// TIA Portal V20 export
DATA_BLOCK "DB_ALARM"   // DB100
{ S7_Optimized_Access := 'FALSE' }
// stored: AutoNumber false
   VAR
      ALARM : Struct
         ALARM_GLOBAL : Bool;   // globální alarm
         HERMA_ERROR : Bool;
         ALARM_2 : Bool;
         ALARM_3 : Bool;
         ALARM_4 : Bool;
         ALARM_5 : Bool;
         air : Bool;   // nedostatečný tlak vzduchu
         ALARM_7 : Bool;
         ALARM_8 : Bool;
         ALARM_9 : Bool;
         ALARM_10 : Bool;
         ALARM_11 : Bool;
         ALARM_12 : Bool;
         ALARM_13 : Bool;
         ALARM_14 : Bool;
         vypadek_safety_karty : Bool;
      END_STRUCT;
      WRONG : Struct
         NENI_INICIALIZACE : Bool;
         WRONG_global : Bool;
         dvere_L_tevreny : Bool;
         dvere_P_otevreny : Bool;
         WRONG_4 : Bool;
         WRONG_5 : Bool;
         WRONG_6 : Bool;
         WRONG_7 : Bool;
         WRONG_8 : Bool;
         WRONG_9 : Bool;
         WRONG_10 : Bool;
         WRONG_11 : Bool;
         WRONG_12 : Bool;
         WRONG_13 : Bool;
         rop_glob_warning : Bool;
         rop_active_autocale : Bool;
      END_STRUCT;
      OP0 : Struct
         ALARM : Struct
            DOOR_ERROR : Bool;
            ALARM_1 : Bool;
            ALARM_2 : Bool;
            ALARM_3 : Bool;
            ALARM_4 : Bool;
            ALARM_5 : Bool;
            ALARM_6 : Bool;
            ALARM_7 : Bool;
            ALARM_8 : Bool;
            ALARM_9 : Bool;
            ALARM_10 : Bool;
            ALARM_11 : Bool;
            ALARM_12 : Bool;
            ALARM_13 : Bool;
            ALARM_14 : Bool;
            ALARM_15 : Bool;
         END_STRUCT;
         WRONG : Struct
            WRONG_0 : Bool;
            WRONG_1 : Bool;
            WRONG_2 : Bool;
            WRONG_3 : Bool;
            WRONG_4 : Bool;
            WRONG_5 : Bool;
            WRONG_6 : Bool;
            WRONG_7 : Bool;
            WRONG_8 : Bool;
            WRONG_9 : Bool;
            WRONG_10 : Bool;
            WRONG_11 : Bool;
            WRONG_12 : Bool;
            WRONG_13 : Bool;
            WRONG_14 : Bool;
            WRONG_15 : Bool;
         END_STRUCT;
         M_0 : Int;
         M_1 : Int;
         M_2 : Int;
         M_3 : Int;
         M_4 : Int;
         M_5 : Int;
         M_6 : Int;
         M_7 : Int;
         M_8 : Int;
         M_9 : Int;
         M_10 : Int;
         M_11 : Int;
         M_12 : Int;
         M_13 : Int;
         M_14 : Int;
         M_15 : Int;
      END_STRUCT;
      OP1 : Struct
         ALARM : Struct
            dvere_1 : Bool;
            ALARM_1 : Bool;
            ALARM_2 : Bool;
            ALARM_3 : Bool;
            ALARM_4 : Bool;
            ALARM_5 : Bool;
            ALARM_6 : Bool;
            hladina_mimo_mez : Bool;
            ALARM_8 : Bool;
            ALARM_9 : Bool;
            ALARM_10 : Bool;
            ALARM_11 : Bool;
            ALARM_12 : Bool;
            ALARM_13 : Bool;
            ALARM_14 : Bool;
            ALARM_15 : Bool;
         END_STRUCT;
         WRONG : Struct
            WRONG_0 : Bool;
            WRONG_1 : Bool;
            WRONG_2 : Bool;
            WRONG_3 : Bool;
            WRONG_4 : Bool;
            WRONG_5 : Bool;
            WRONG_6 : Bool;
            WRONG_7 : Bool;
            WRONG_8 : Bool;
            WRONG_9 : Bool;
            WRONG_10 : Bool;
            WRONG_11 : Bool;
            WRONG_12 : Bool;
            WRONG_13 : Bool;
            WRONG_14 : Bool;
            WRONG_15 : Bool;
         END_STRUCT;
         "-Y7_KARUSEL" : Int;
         "-Y9_ZARAZKA" : Int;
         M_2 : Int;
         M_3 : Int;
         M_4 : Int;
         M_5 : Int;
         M_6 : Int;
         M_7 : Int;
         M_8 : Int;
         M_9 : Int;
         M_10 : Int;
         M_11 : Int;
         M_12 : Int;
         M_13 : Int;
         M_14 : Int;
         M_15 : Int;
      END_STRUCT;
      OP2 : Struct
         ALARM : Struct
            dvere_1 : Bool;
            dvere_2 : Bool;
            dvere_3 : Bool;
            dvere_4 : Bool;
            paprsek : Bool;
            porucha_svarovani : Bool;
            rop_alarm : Bool;
            servo_power_error : Bool;
            servo_jog_error : Bool;
            servo_homing : Bool;
            Cel_podel_porucha : Bool;
            vysoka_tuzka : Bool;
            ALARM_12 : Bool;
            ALARM_13 : Bool;
            folie : Bool;
            ALARM_15 : Bool;
         END_STRUCT;
         WRONG : Struct
            WRONG_0 : Bool;
            WRONG_1 : Bool;
            WRONG_2 : Bool;
            WRONG_3 : Bool;
            WRONG_4 : Bool;
            WRONG_5 : Bool;
            WRONG_6 : Bool;
            WRONG_7 : Bool;
            WRONG_8 : Bool;
            WRONG_9 : Bool;
            WRONG_10 : Bool;
            WRONG_11 : Bool;
            WRONG_12 : Bool;
            WRONG_13 : Bool;
            WRONG_14 : Bool;
            WRONG_15 : Bool;
         END_STRUCT;
         A1 : Int;   // -YA1
         A2 : Int;   // -YA2
         A3 : Int;   // -YA3
         A4 : Int;   // -YA4
         A5 : Int;   // -YA5
         A6 : Int;   // -YA6
         A7 : Int;   // -YA7
         A8 : Int;   // -YA8
         M_8 : Int;
         M_9 : Int;
         M_10 : Int;
         M_11 : Int;
         M_12 : Int;
         M_13 : Int;
         M_14 : Int;
         M_15 : Int;
      END_STRUCT;
      OP3 : Struct
         ALARM : Struct
            ALARM_0 : Bool;
            ALARM_1 : Bool;
            ALARM_2 : Bool;
            ALARM_3 : Bool;
            ALARM_4 : Bool;
            ALARM_5 : Bool;
            ALARM_6 : Bool;
            ALARM_7 : Bool;
            ALARM_8 : Bool;
            ALARM_9 : Bool;
            ALARM_10 : Bool;
            ALARM_11 : Bool;
            ALARM_12 : Bool;
            ALARM_13 : Bool;
            ALARM_14 : Bool;
            ALARM_15 : Bool;
         END_STRUCT;
         WRONG : Struct
            WRONG_0 : Bool;
            WRONG_1 : Bool;
            WRONG_2 : Bool;
            WRONG_3 : Bool;
            WRONG_4 : Bool;
            WRONG_5 : Bool;
            WRONG_6 : Bool;
            WRONG_7 : Bool;
            WRONG_8 : Bool;
            WRONG_9 : Bool;
            WRONG_10 : Bool;
            WRONG_11 : Bool;
            WRONG_12 : Bool;
            WRONG_13 : Bool;
            WRONG_14 : Bool;
            WRONG_15 : Bool;
         END_STRUCT;
         B1 : Int;   // -YB1
         B2 : Int;   // -YB2
         B3 : Int;   // -YB3
         B4 : Int;   // -YB4
         B5 : Int;   // -YB5
         B6 : Int;   // -YB6
         B7 : Int;   // -YB7
         B8 : Int;   // -YB8
         M_8 : Int;
         M_9 : Int;
         M_10 : Int;
         M_11 : Int;
         M_12 : Int;
         M_13 : Int;
         M_14 : Int;
         M_15 : Int;
      END_STRUCT;
      OP4 : Struct
         ALARM : Struct
            odsavani_nefunguje : Bool;
            ALARM_1 : Bool;
            ALARM_2 : Bool;
            ALARM_3 : Bool;
            ALARM_4 : Bool;
            ALARM_5 : Bool;
            ALARM_6 : Bool;
            ALARM_7 : Bool;
            ALARM_8 : Bool;
            ALARM_9 : Bool;
            ALARM_10 : Bool;
            ALARM_11 : Bool;
            ALARM_12 : Bool;
            ALARM_13 : Bool;
            ALARM_14 : Bool;
            ALARM_15 : Bool;
         END_STRUCT;
         WRONG : Struct
            WRONG_0 : Bool;
            WRONG_1 : Bool;
            WRONG_2 : Bool;
            WRONG_3 : Bool;
            WRONG_4 : Bool;
            WRONG_5 : Bool;
            WRONG_6 : Bool;
            WRONG_7 : Bool;
            WRONG_8 : Bool;
            WRONG_9 : Bool;
            WRONG_10 : Bool;
            WRONG_11 : Bool;
            WRONG_12 : Bool;
            WRONG_13 : Bool;
            WRONG_14 : Bool;
            WRONG_15 : Bool;
         END_STRUCT;
         M_0 : Int;
         M_1 : Int;
         M_2 : Int;
         M_3 : Int;
         M_4 : Int;
         M_5 : Int;
         M_6 : Int;
         M_7 : Int;
         M_8 : Int;
         M_9 : Int;
         M_10 : Int;
         M_11 : Int;
         M_12 : Int;
         M_13 : Int;
         M_14 : Int;
         M_15 : Int;
      END_STRUCT;
      OP5 : Struct
         ALARM : Struct
            ALARM_0 : Bool;
            ALARM_1 : Bool;
            ALARM_2 : Bool;
            ALARM_3 : Bool;
            ALARM_4 : Bool;
            ALARM_5 : Bool;
            ALARM_6 : Bool;
            ALARM_7 : Bool;
            ALARM_8 : Bool;
            ALARM_9 : Bool;
            ALARM_10 : Bool;
            ALARM_11 : Bool;
            ALARM_12 : Bool;
            ALARM_13 : Bool;
            ALARM_14 : Bool;
            ALARM_15 : Bool;
         END_STRUCT;
         WRONG : Struct
            WRONG_0 : Bool;
            WRONG_1 : Bool;
            WRONG_2 : Bool;
            WRONG_3 : Bool;
            WRONG_4 : Bool;
            WRONG_5 : Bool;
            WRONG_6 : Bool;
            WRONG_7 : Bool;
            WRONG_8 : Bool;
            WRONG_9 : Bool;
            WRONG_10 : Bool;
            WRONG_11 : Bool;
            WRONG_12 : Bool;
            WRONG_13 : Bool;
            WRONG_14 : Bool;
            WRONG_15 : Bool;
         END_STRUCT;
         M_0 : Int;
         M_1 : Int;
         M_2 : Int;
         M_3 : Int;
         M_4 : Int;
         M_5 : Int;
         M_6 : Int;
         M_7 : Int;
         M_8 : Int;
         M_9 : Int;
         M_10 : Int;
         M_11 : Int;
         M_12 : Int;
         M_13 : Int;
         M_14 : Int;
         M_15 : Int;
      END_STRUCT;
      null : Struct
         ALARM_0 : Bool;
         ALARM_1 : Bool;
         ALARM_2 : Bool;
         ALARM_3 : Bool;
         ALARM_4 : Bool;
         ALARM_5 : Bool;
         ALARM_6 : Bool;
         ALARM_7 : Bool;
         ALARM_8 : Bool;
         ALARM_9 : Bool;
         ALARM_10 : Bool;
         ALARM_11 : Bool;
         ALARM_12 : Bool;
         ALARM_13 : Bool;
         ALARM_14 : Bool;
         ALARM_15 : Bool;
      END_STRUCT;
      alarmy : Array[0..255] of Bool;
      alarm_line : Int;
      wrong_line : Int;
      alarm_op_1 : Int;
      wrong_op_1 : Int;
      alarm_op_2 : Int;
      wrong_op_2 : Int;
      alarm_op_3 : Int;
      wrong_op_3 : Int;
      alarm_op_4 : Int;
      wrong_op_4 : Int;
      alarm_op_5 : Int;
      wrong_op_5 : Int;
      T_tiskarna : TON_TIME;
   END_VAR
BEGIN
END_DATA_BLOCK
